(* IEC 61131-3 sources: volt/packages/volt-lsp-iec/test-corpus/pro2193/Device/Plc Logic/Application/09 Misc/Library Manager/OMAC_PackML_State_Machine, 7 files *)

(* ---- STATE.dut ---- *)
TYPE STATE :
(
	STOPPED := 16#1,
	RESETTING := 16#2,
	IDLE := 16#4,
	STARTING := 16#8,
	EXECUTE := 16#10,
	HOLDING := 16#20,
	HELD := 16#40,
	UNHOLDING := 16#80,
	SUSPENDING := 16#100,
	SUSPENDED := 16#200,
	UNSUSPENDING := 16#400,
	COMPLETING := 16#800,
	COMPLETE := 16#1000,
	STOPPING := 16#2000,
	ABORTING := 16#4000,
	ABORTED := 16#8000,
	CLEARING := 16#10000,
	NO := 0,
	ALL := 16#1FFFF,
	INVALID := 16#80000000
);
END_TYPE

(* ---- GVL.gvl ---- *)
VAR_GLOBAL
	GC_USIMAXMODES : USINT := 10;
END_VAR

(* ---- IUNITMODE.itf ---- *)
INTERFACE IUNITMODE
END_INTERFACE

METHOD ABORT : BOOL
END_METHOD

METHOD ACTINGSTATECOMPLETED : BOOL
END_METHOD

METHOD CLEAR : BOOL
END_METHOD

METHOD HOLD : BOOL
END_METHOD

METHOD RESET : BOOL
END_METHOD

METHOD START : BOOL
END_METHOD

METHOD STOP : BOOL
END_METHOD

METHOD SUSPEND : BOOL
END_METHOD

METHOD UNHOLD : BOOL
END_METHOD

METHOD UNSUSPEND : BOOL
END_METHOD

METHOD ALLOWSENTERING : BOOL
VAR_INPUT
	E : State;
END_VAR
END_METHOD

METHOD ENTER : BOOL
VAR_INPUT
	E : State;
END_VAR
END_METHOD

METHOD NEXTSTATE : State
VAR_INPUT
	E : State;
END_VAR
END_METHOD

(* ---- GLOBALTEXTLIST.pou ---- *)
FUNCTION_BLOCK GLOBALTEXTLIST
VAR
	M_TEXTLISTFILE : STRING(255);
	_STNAMESPACE : STRING;
END_VAR
END_FUNCTION_BLOCK

(* ---- IMAGEPOOL.pou ---- *)
FUNCTION_BLOCK IMAGEPOOL
VAR
	M_STNAMESPACE : STRING(80);
	M_STHELPVARID : STRING;
	M_STHELPVARPATH : STRING(255);
	M_STHELP : STRING;
	M_REGISTERIMAGES : BOOL := TRUE;
END_VAR
END_FUNCTION_BLOCK

METHOD FB_INIT : BOOL
VAR_INPUT
	BINITRETAINS : BOOL;
	BINCOPYCODE : BOOL;
END_VAR
END_METHOD

METHOD FB_REINIT : BOOL
END_METHOD

METHOD FB_EXIT : BOOL
VAR_INPUT
	BINCOPYCODE : BOOL;
END_VAR
END_METHOD

(* ---- UNITMODE.pou ---- *)
FUNCTION_BLOCK UNITMODE
VAR_INPUT
	SNAME : STRING;
	DWSUPPORTEDSTATES : DWORD := 2#11111111111111111;
	DWALLOWSLEAVINGFROMSTATES : DWORD := (State.Stopped OR State.Aborted);
	DWALLOWSENTERINGINTOSTATES : DWORD := (State.Stopped OR State.Aborted);
	EINITIALSTATE : State;
	XACTIVE : BOOL;
END_VAR
VAR
	ESTATE : State := State.Invalid;
	BINIT : BOOL;
	ACTIVE : BOOL;
	ALLOWSLEAVING : BOOL;
	CURRENTSTATE : State;
	NAME : STRING;
	SUPPORTEDSTATES : DWORD;
END_VAR
END_FUNCTION_BLOCK

METHOD ABORT : BOOL
END_METHOD

METHOD ACTINGSTATECOMPLETED : BOOL
END_METHOD

METHOD CLEAR : BOOL
END_METHOD

METHOD HOLD : BOOL
END_METHOD

METHOD RESET : BOOL
END_METHOD

METHOD START : BOOL
END_METHOD

METHOD STOP : BOOL
END_METHOD

METHOD SUSPEND : BOOL
END_METHOD

METHOD UNHOLD : BOOL
END_METHOD

METHOD UNSUSPEND : BOOL
END_METHOD

METHOD ALLOWSENTERING : BOOL
VAR_INPUT
	E : State;
END_VAR
END_METHOD

METHOD ENTER : BOOL
VAR_INPUT
	E : State;
END_VAR
END_METHOD

METHOD NEXTSTATE : State
VAR_INPUT
	E : State;
END_VAR
END_METHOD

(* ---- UNITMODEMANAGER.pou ---- *)
FUNCTION_BLOCK UNITMODEMANAGER
VAR
	APUM : ARRAY [1..gc_usiMaxModes] OF IUnitMode;
	USINUMBEROFUMS : USINT := 0;
	USIACTUALUM : USINT;
	ACTIVEUNITMODE : IUnitMode;
	ACTIVEUNITMODENUMBER : USINT;
END_VAR
END_FUNCTION_BLOCK

METHOD ALLOWSSWITCHINGTO : BOOL
VAR_INPUT
	USI : USINT;
END_VAR
END_METHOD

METHOD FINDMODE : USINT
VAR_INPUT
	SNAME : STRING;
END_VAR
END_METHOD

METHOD REGISTER : BOOL
VAR_INPUT
	PUM : IUnitMode;
END_VAR
END_METHOD

METHOD SWITCHUNITMODE : BOOL
VAR_INPUT
	SNEWMODENAME : STRING;
END_VAR
END_METHOD
